(* IEC 61131-3 sources: plc-vscode/tests/st/test-ready/rusty/libs/stdlib/iec61131-st (part 3) *)

(* ---- counters.st ---- *)
(******************************************************************************
Description: Counter up
Input:
  - CU: Count up
  - R: Reset counter to 0
  - PV: Counter limit
Output:
  - Q: Counter reached limit
  - CV: Current counter value
Return: Output is used as return value
******************************************************************************)
{external}
FUNCTION_BLOCK CTU
VAR_INPUT
    CU : BOOL;
    R : BOOL;
    PV : INT;
END_VAR
VAR_OUTPUT
    Q : BOOL;
    CV : INT;
END_VAR
VAR
    M : BOOL;
END_VAR
END_FUNCTION_BLOCK

(******************************************************************************
Description: Counter up
Input:
  - CU: Count up
  - R: Reset counter to 0
  - PV: Counter limit
Output:
  - Q: Counter reached limit
  - CV: Current counter value
Return: Output is used as return value
******************************************************************************)
{external}
FUNCTION_BLOCK CTU_INT
VAR_INPUT
    CU : BOOL;
    R : BOOL;
    PV : INT;
END_VAR
VAR_OUTPUT
    Q : BOOL;
    CV : INT;
END_VAR
VAR
    M : BOOL;
END_VAR
END_FUNCTION_BLOCK

(******************************************************************************
Description: Counter up
Input:
  - CU: Count up
  - R: Reset counter to 0
  - PV: Counter limit
Output:
  - Q: Counter reached limit
  - CV: Current counter value
Return: Output is used as return value
******************************************************************************)
{external}
FUNCTION_BLOCK CTU_DINT
VAR_INPUT
    CU : BOOL;
    R : BOOL;
    PV : DINT;
END_VAR
VAR_OUTPUT
    Q : BOOL;
    CV : DINT;
END_VAR
VAR
    M : BOOL;
END_VAR
END_FUNCTION_BLOCK

(******************************************************************************
Description: Counter up
Input:
  - CU: Count up
  - R: Reset counter to 0
  - PV: Counter limit
Output:
  - Q: Counter reached limit
  - CV: Current counter value
Return: Output is used as return value
******************************************************************************)
{external}
FUNCTION_BLOCK CTU_UDINT
VAR_INPUT
    CU : BOOL;
    R : BOOL;
    PV : UDINT;
END_VAR
VAR_OUTPUT
    Q : BOOL;
    CV : UDINT;
END_VAR
VAR
    M : BOOL;
END_VAR
END_FUNCTION_BLOCK

(******************************************************************************
Description: Counter up
Input:
  - CU: Count up
  - R: Reset counter to 0
  - PV: Counter limit
Output:
  - Q: Counter reached limit
  - CV: Current counter value
Return: Output is used as return value
******************************************************************************)
{external}
FUNCTION_BLOCK CTU_LINT
VAR_INPUT
    CU : BOOL;
    R : BOOL;
    PV : LINT;
END_VAR
VAR_OUTPUT
    Q : BOOL;
    CV : LINT;
END_VAR
VAR
    M : BOOL;
END_VAR
END_FUNCTION_BLOCK

(******************************************************************************
Description: Counter up
Input:
  - CU: Count up
  - R: Reset counter to 0
  - PV: Counter limit
Output:
  - Q: Counter reached limit
  - CV: Current counter value
Return: Output is used as return value
******************************************************************************)
{external}
FUNCTION_BLOCK CTU_ULINT
VAR_INPUT
    CU : BOOL;
    R : BOOL;
    PV : ULINT;
END_VAR
VAR_OUTPUT
    Q : BOOL;
    CV : ULINT;
END_VAR
VAR
    M : BOOL;
END_VAR
END_FUNCTION_BLOCK

(******************************************************************************
Description: Counter down
Input:
  - CD: Count down
  - LD: Load start value
  - PV: Start value
Output:
  - Q: Counter reached 0
  - CV: Current counter value
Return: Output is used as return value
******************************************************************************)
{external}
FUNCTION_BLOCK CTD
VAR_INPUT
    CD : BOOL;
    LD : BOOL;
    PV : INT;
END_VAR
VAR_OUTPUT
    Q : BOOL;
    CV : INT;
END_VAR
VAR
    M : BOOL;
END_VAR
END_FUNCTION_BLOCK

(******************************************************************************
Description: Counter down
Input:
  - CD: Count down
  - LD: Load start value
  - PV: Start value
Output:
  - Q: Counter reached 0
  - CV: Current counter value
Return: Output is used as return value
******************************************************************************)
{external}
FUNCTION_BLOCK CTD_INT
VAR_INPUT
    CD : BOOL;
    LD : BOOL;
    PV : INT;
END_VAR
VAR_OUTPUT
    Q : BOOL;
    CV : INT;
END_VAR
VAR
    M : BOOL;
END_VAR
END_FUNCTION_BLOCK

(******************************************************************************
Description: Counter down
Input:
  - CD: Count down
  - LD: Load start value
  - PV: Start value
Output:
  - Q: Counter reached 0
  - CV: Current counter value
Return: Output is used as return value
******************************************************************************)
{external}
FUNCTION_BLOCK CTD_DINT
VAR_INPUT
    CD : BOOL;
    LD : BOOL;
    PV : DINT;
END_VAR
VAR_OUTPUT
    Q : BOOL;
    CV : DINT;
END_VAR
VAR
    M : BOOL;
END_VAR
END_FUNCTION_BLOCK

(******************************************************************************
Description: Counter down
Input:
  - CD: Count down
  - LD: Load start value
  - PV: Start value
Output:
  - Q: Counter reached 0
  - CV: Current counter value
Return: Output is used as return value
******************************************************************************)
{external}
FUNCTION_BLOCK CTD_UDINT
VAR_INPUT
    CD : BOOL;
    LD : BOOL;
    PV : UDINT;
END_VAR
VAR_OUTPUT
    Q : BOOL;
    CV : UDINT;
END_VAR
VAR
    M : BOOL;
END_VAR
END_FUNCTION_BLOCK

(******************************************************************************
Description: Counter down
Input:
  - CD: Count down
  - LD: Load start value
  - PV: Start value
Output:
  - Q: Counter reached 0
  - CV: Current counter value
Return: Output is used as return value
******************************************************************************)
{external}
FUNCTION_BLOCK CTD_LINT
VAR_INPUT
    CD : BOOL;
    LD : BOOL;
    PV : LINT;
END_VAR
VAR_OUTPUT
    Q : BOOL;
    CV : LINT;
END_VAR
VAR
    M : BOOL;
END_VAR
END_FUNCTION_BLOCK

(******************************************************************************
Description: Counter down
Input:
  - CD: Count down
  - LD: Load start value
  - PV: Start value
Output:
  - Q: Counter reached 0
  - CV: Current counter value
Return: Output is used as return value
******************************************************************************)
{external}
FUNCTION_BLOCK CTD_ULINT
VAR_INPUT
    CD : BOOL;
    LD : BOOL;
    PV : ULINT;
END_VAR
VAR_OUTPUT
    Q : BOOL;
    CV : ULINT;
END_VAR
VAR
    M : BOOL;
END_VAR
END_FUNCTION_BLOCK

(******************************************************************************
Description: Counter up and down
Input:
  - CU: Count up
  - CD: Count down
  - R: Reset counter to 0
  - LD: Load start value
  - PV: Start value / counter limit
Output:
  - QU: Counter reached limit
  - QD: Counter reached  0
  - CV: Current counter value
Return: Output is used as return value
******************************************************************************)
{external}
FUNCTION_BLOCK CTUD
VAR_INPUT
    CU : BOOL;
    CD : BOOL;
    R : BOOL;
    LD : BOOL;
    PV : INT;
END_VAR
VAR_OUTPUT
    QU : BOOL;
    QD : BOOL;
    CV : INT;
END_VAR
VAR
    MU : BOOL;
    MD : BOOL;
END_VAR
END_FUNCTION_BLOCK

(******************************************************************************
Description: Counter up and down
Input:
  - CU: Count up
  - CD: Count down
  - R: Reset counter to 0
  - LD: Load start value
  - PV: Start value / counter limit
Output:
  - QU: Counter reached limit
  - QD: Counter reached  0
  - CV: Current counter value
Return: Output is used as return value
******************************************************************************)
{external}
FUNCTION_BLOCK CTUD_INT
VAR_INPUT
    CU : BOOL;
    CD : BOOL;
    R : BOOL;
    LD : BOOL;
    PV : INT;
END_VAR
VAR_OUTPUT
    QU : BOOL;
    QD : BOOL;
    CV : INT;
END_VAR
VAR
    MU : BOOL;
    MD : BOOL;
END_VAR
END_FUNCTION_BLOCK

(******************************************************************************
Description: Counter up and down
Input:
  - CU: Count up
  - CD: Count down
  - R: Reset counter to 0
  - LD: Load start value
  - PV: Start value / counter limit
Output:
  - QU: Counter reached limit
  - QD: Counter reached  0
  - CV: Current counter value
Return: Output is used as return value
******************************************************************************)
{external}
FUNCTION_BLOCK CTUD_DINT
VAR_INPUT
    CU : BOOL;
    CD : BOOL;
    R : BOOL;
    LD : BOOL;
    PV : DINT;
END_VAR
VAR_OUTPUT
    QU : BOOL;
    QD : BOOL;
    CV : DINT;
END_VAR
VAR
    MU : BOOL;
    MD : BOOL;
END_VAR
END_FUNCTION_BLOCK

(******************************************************************************
Description: Counter up and down
Input:
  - CU: Count up
  - CD: Count down
  - R: Reset counter to 0
  - LD: Load start value
  - PV: Start value / counter limit
Output:
  - QU: Counter reached limit
  - QD: Counter reached  0
  - CV: Current counter value
Return: Output is used as return value
******************************************************************************)
{external}
FUNCTION_BLOCK CTUD_UDINT
VAR_INPUT
    CU : BOOL;
    CD : BOOL;
    R : BOOL;
    LD : BOOL;
    PV : UDINT;
END_VAR
VAR_OUTPUT
    QU : BOOL;
    QD : BOOL;
    CV : UDINT;
END_VAR
VAR
    MU : BOOL;
    MD : BOOL;
END_VAR
END_FUNCTION_BLOCK

(******************************************************************************
Description: Counter up and down
Input:
  - CU: Count up
  - CD: Count down
  - R: Reset counter to 0
  - LD: Load start value
  - PV: Start value / counter limit
Output:
  - QU: Counter reached limit
  - QD: Counter reached  0
  - CV: Current counter value
Return: Output is used as return value
******************************************************************************)
{external}
FUNCTION_BLOCK CTUD_LINT
VAR_INPUT
    CU : BOOL;
    CD : BOOL;
    R : BOOL;
    LD : BOOL;
    PV : LINT;
END_VAR
VAR_OUTPUT
    QU : BOOL;
    QD : BOOL;
    CV : LINT;
END_VAR
VAR
    MU : BOOL;
    MD : BOOL;
END_VAR
END_FUNCTION_BLOCK

(******************************************************************************
Description: Counter up and down
Input:
  - CU: Count up
  - CD: Count down
  - R: Reset counter to 0
  - LD: Load start value
  - PV: Start value / counter limit
Output:
  - QU: Counter reached limit
  - QD: Counter reached  0
  - CV: Current counter value
Return: Output is used as return value
******************************************************************************)
{external}
FUNCTION_BLOCK CTUD_ULINT
VAR_INPUT
    CU : BOOL;
    CD : BOOL;
    R : BOOL;
    LD : BOOL;
    PV : ULINT;
END_VAR
VAR_OUTPUT
    QU : BOOL;
    QD : BOOL;
    CV : ULINT;
END_VAR
VAR
    MU : BOOL;
    MD : BOOL;
END_VAR
END_FUNCTION_BLOCK

(* ---- flanks.st ---- *)
(******************************************************************************
Description: Rising Edge detection
Input:
  - CLK:  Signal to detect
Output:
  - Q:  Edge detected
Return: Output variable are used for return.
******************************************************************************)
{external}
FUNCTION_BLOCK R_TRIG
VAR_INPUT
    CLK: BOOL;
END_VAR
VAR_OUTPUT
    Q: BOOL;
END_VAR
VAR
    M: BOOL;
END_VAR
END_FUNCTION_BLOCK

(******************************************************************************
Description: Falling Edge detection
Input:
  - CLK:  Signal to detect
Output:
  - Q:  Edge detected
Return: Output variable is used for return.
******************************************************************************)
{external}
FUNCTION_BLOCK F_TRIG
VAR_INPUT
    CLK: BOOL;
END_VAR
VAR_OUTPUT
    Q: BOOL;
END_VAR
VAR
    M: BOOL;
END_VAR
END_FUNCTION_BLOCK

(* ---- timers.st ---- *)
{external}
(******************************************************************************
Description: Timer Pulse
Input:
  - IN: Trigger for Start of the Signal
  - PT: The length of the High-Signal
Output:
  - Q: The pulse
  - ET: The current phase of the High-Signal
Return: Output variables are used for return.
******************************************************************************)
FUNCTION_BLOCK TP
    VAR_INPUT
        IN : BOOL;
        PT : TIME;
    END_VAR
    VAR_OUTPUT
        Q  : BOOL;
        ET : TIME;
    END_VAR
    VAR
        __signal__ : BOOL; (* Value representing the internal signal *)
        __is_running__: BOOL; (* Internal flag to track timer on/off state *)
        __BUFFER__ : ARRAY[1..24] OF BYTE; (* Buffer used for internal implementation *)
    END_VAR
END_FUNCTION_BLOCK

{external}
(******************************************************************************
Description: Timer Pulse
Input:
  - IN: Trigger for Start of the Signal
  - PT: The length of the High-Signal
Output:
  - Q: The pulse
  - ET: The current phase of the High-Signal
Return: Output variables are used for return.
******************************************************************************)
FUNCTION_BLOCK TP_TIME
    VAR_INPUT
        IN : BOOL;
        PT : TIME;
    END_VAR
    VAR_OUTPUT
        Q  : BOOL;
        ET : TIME;
    END_VAR
    VAR
      __signal__ : BOOL; (* Value representing the internal signal *)
      __is_running__: BOOL; (* Internal flag to track timer on/off state *)
      __BUFFER__ : ARRAY[1..24] OF BYTE; (* Buffer used for internal implementation *)
    END_VAR
END_FUNCTION_BLOCK

{external}
(******************************************************************************
Description: Timer Pulse
Input:
  - IN: Trigger for Start of the Signal
  - PT: The length of the High-Signal
Output:
  - Q: The pulse
  - ET: The current phase of the High-Signal
Return: Output variables are used for return.
******************************************************************************)
FUNCTION_BLOCK TP_LTIME
    VAR_INPUT
        IN : BOOL;
        PT : TIME;
    END_VAR
    VAR_OUTPUT
        Q  : BOOL;
        ET : LTIME;
    END_VAR
    VAR
        __signal__ : BOOL; (* Value representing the internal signal *)
        __is_running__: BOOL; (* Internal flag to track timer on/off state *)
        __BUFFER__ : ARRAY[1..24] OF BYTE; (* Buffer used for internal implementation *)
    END_VAR
END_FUNCTION_BLOCK

{external}
(******************************************************************************
Description: Timer on delay.
Input:
  - IN: Starts timer with rising edge, resets timer with falling edge
  - PT: Time to pass, before Q is set
Output:
  - Q: Is TRUE, PT seconds after IN had a rising edge
  - ET: Elapsed time
Return: Output variables are used for return.
******************************************************************************)
FUNCTION_BLOCK TON
VAR_INPUT
    IN: BOOL;
    PT: TIME;
END_VAR
VAR_OUTPUT
    Q: BOOL;
    ET: TIME;
END_VAR
VAR
  __signal__ : BOOL; (* Value representing the internal signal *)
  __is_running__: BOOL; (* Internal flag to track timer on/off state *)
  __BUFFER__ : ARRAY[1..24] OF BYTE; (* Buffer used for internal implementation *)
END_VAR
END_FUNCTION_BLOCK

{external}
(******************************************************************************
Description: Timer on delay.
Input:
  - IN: Starts timer with rising edge, resets timer with falling edge
  - PT: Time to pass, before Q is set
Output:
  - Q: Is TRUE, PT seconds after IN had a rising edge
  - ET: Elapsed time
Return: Output variables are used for return.
******************************************************************************)
FUNCTION_BLOCK TON_TIME
VAR_INPUT
    IN: BOOL;
    PT: TIME;
END_VAR
VAR_OUTPUT
    Q: BOOL;
    ET: TIME;
END_VAR
VAR
  __signal__ : BOOL; (* Value representing the internal signal *)
  __is_running__: BOOL; (* Internal flag to track timer on/off state *)
  __BUFFER__ : ARRAY[1..24] OF BYTE; (* Buffer used for internal implementation *)
END_VAR
END_FUNCTION_BLOCK

{external}
(******************************************************************************
Description: Timer on delay.
Input:
  - IN: Starts timer with rising edge, resets timer with falling edge
  - PT: Time to pass, before Q is set
Output:
  - Q: Is TRUE, PT seconds after IN had a rising edge
  - ET: Elapsed time
Return: Output variables are used for return.
******************************************************************************)
FUNCTION_BLOCK TON_LTIME
VAR_INPUT
    IN: BOOL;
    PT: LTIME;
END_VAR
VAR_OUTPUT
    Q: BOOL;
    ET: TIME;
END_VAR
VAR
  __signal__ : BOOL; (* Value representing the internal signal *)
  __is_running__: BOOL; (* Internal flag to track timer on/off state *)
  __BUFFER__ : ARRAY[1..24] OF BYTE; (* Buffer used for internal implementation *)
END_VAR
END_FUNCTION_BLOCK

{external}
(******************************************************************************
Description: Timer of delay
Input:
  - IN: Starts timer with falling edge, resets timer with rising edge
  - PT: Time to pass, before Q is set
Output:
  - Q: is FALSE, PT seconds after IN had a falling edge
  - ET: Elapsed time
Return: Output variables are used for return.
******************************************************************************)
FUNCTION_BLOCK TOF
VAR_INPUT
    IN: BOOL;
    PT:TIME;
END_VAR
VAR_OUTPUT
    Q: BOOL;
    ET: TIME;
END_VAR
VAR
  __signal__ : BOOL; (* Value representing the internal signal *)
  __is_running__: BOOL; (* Internal flag to track timer on/off state *)
  __BUFFER__ : ARRAY[1..24] OF BYTE; (* Buffer used for internal implementation *)
END_VAR
END_FUNCTION_BLOCK

{external}
(******************************************************************************
Description: Timer of delay
Input:
  - IN: Starts timer with falling edge, resets timer with rising edge
  - PT: Time to pass, before Q is set
Output:
  - Q: is FALSE, PT seconds after IN had a falling edge
  - ET: Elapsed time
Return: Output variables are used for return.
******************************************************************************)
FUNCTION_BLOCK TOF_TIME
VAR_INPUT
    IN: BOOL;
    PT:TIME;
END_VAR
VAR_OUTPUT
    Q: BOOL;
    ET: TIME;
END_VAR
VAR
  __signal__ : BOOL; (* Value representing the internal signal *)
  __is_running__: BOOL; (* Internal flag to track timer on/off state *)
  __BUFFER__ : ARRAY[1..24] OF BYTE; (* Buffer used for internal implementation *)
END_VAR
END_FUNCTION_BLOCK

{external}
(******************************************************************************
Description: Timer of delay
Input:
  - IN: Starts timer with falling edge, resets timer with rising edge
  - PT: Time to pass, before Q is set
Output:
  - Q: is FALSE, PT seconds after IN had a falling edge
  - ET: Elapsed time
Return: Output variables are used for return.
******************************************************************************)
FUNCTION_BLOCK TOF_LTIME
VAR_INPUT
    IN: BOOL;
    PT:LTIME;
END_VAR
VAR_OUTPUT
    Q: BOOL;
    ET: LTIME;
END_VAR
VAR
  __signal__ : BOOL; (* Value representing the internal signal *)
  __is_running__: BOOL; (* Internal flag to track timer on/off state *)
  __BUFFER__ : ARRAY[1..24] OF BYTE; (* Buffer used for internal implementation *)
END_VAR
END_FUNCTION_BLOCK
